(* Buzzer Sounds on Fault or Completion *)

PROGRAM main
  VAR
    InputA AT %MX0.1 : BOOL;
    InputB AT %MX0.2 : BOOL;
    Output AT %QX0.1 : BOOL; (* Output Buzzer *)
  END_VAR

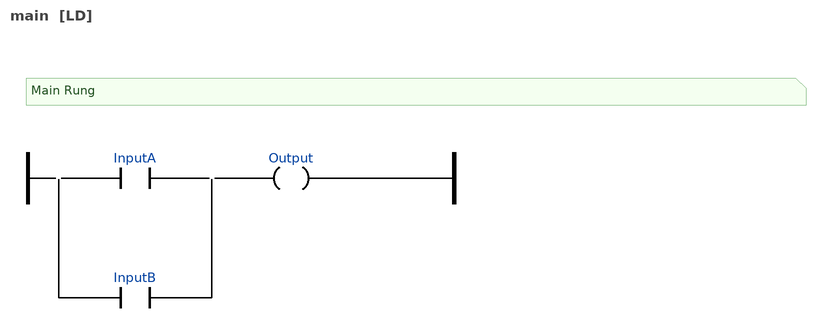
(* LD diagram, written out as Structured Text *)
(* Main Rung *)
Output := InputA OR InputB;
END_PROGRAM
